Fanuc KAREL source: kt00092.KL

-- PROVISIONAL review KL for V770-1; original PC SHA256 cda63a8d707f777b41503394bcfb93cb2d058fa61a209636ded42372794e6350
-- Incomplete behavior may be omitted. Consult companion uncertainty JSON. Do not deploy.
PROGRAM KT00092
%NOLOCKGROUP
VAR
  R2 : REAL
  OUT : REAL
-- UNRESOLVED_DECL H1 type=002017
BEGIN
  -- UNRESOLVED_PC offsets 5-19; opcodes 2E,22,9D,33,B4
  -- UNRESOLVED_PC offsets 24-35; opcodes 2E,23
  -- UNRESOLVED_PC offsets 40-64; opcodes 22,9D,33,B3,21,29,64,6B,23
  -- UNRESOLVED_PC offsets 69-73; opcodes 7F
END KT00092
